SUBAPPLICATION Button_Toggle_RPC_TO_Remote_BG_Option_OPC (* Wie Button_Toggle_RPC_TO_Remote_BG_OPC (IO-Diag-Taster, Loslassen ruft per CLIENT_0 eine RPC-Toggle-Methode auf dem Zielmodul auf, Hintergrundfarbe aus Remote-Subscribe), aber per AOption aktiviert statt QI/INIT. AOption_OUT reicht die Aktivierung nach dem eigenen INIT weiter (Daisy-Chain). *)
  (* Standard: 61499-2; Description: Copyright (c) 2026 Meisterschulen am Ostbahnhof This program and the accompanying materials are made available under the terms of the Eclipse Public License 2.0 which is available at https://www.eclipse.org/legal/epl-2.0/ SPDX-License-Identifier: EPL-2.0 *)
  (* Version 1.1, 2026-10-30, Franz Höpfinger, Meisterschulen am Ostbahnhof, Remote-Clients mit Remote_Init_Retry: Kette (und Option-INIT_CNF) wartet nicht mehr auf die Gegenstation, nach INITO- neuer Versuch nach 2 s (forte #1092, sonst 60 s pro fehlendem Node und danach tot). *)
  (* Version 1.0, 2026-10-17, Franz Höpfinger, Meisterschulen am Ostbahnhof, Kopie von Button_Toggle_RPC_TO_Remote_BG_OPC (Franz: 'kopieren, Variante mit AOption machen') - INIT/INITO/QI/QO ersetzt durch AOption_IN (AOption_X_TO_EVENT) und AOption_OUT (AOption_EVENT_TO_X, Daisy-Chain wie OptionalGroup_001a). AOption_OUT muss weiterverbunden sein (DummyGroup als Kettenende), sonst kommt kein INIT_CNF zurueck. *)
  PACKAGE MyLib::sys;
  IMPORT isobus::UT::Q::const::IDs::ID_NULL;
  IMPORT isobus::UT::io::Button::ButtonActivationCode::BT_RELEASED_UNLATCHED;
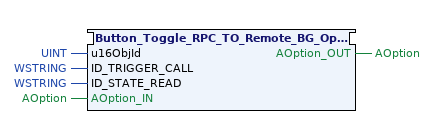
  VAR_INPUT
    u16ObjId : UINT := ID_NULL; (* Object ID Button/Background *)
    ID_TRIGGER_CALL : WSTRING; (* Remote-Methodenadresse (ACTION=CALL_METHOD) fuer den argumentlosen Trigger-Methodenaufruf auf dem Zielmodul *)
    ID_STATE_READ : WSTRING; (* Lokal ueberwachte Adresse (BOOL, ACTION=READ) fuer den Flipflop-Zustand, wird vom Zielmodul remote beschrieben *)
  END_VAR
  SOCKETS
    AOption_IN : Option::AOption; (* Treibt INIT/QI - anschliessen an AOption_AUI_DEMUX_N.OUTx oder AOption_OUT einer vorgeschalteten Instanz *)
  END_SOCKETS
  PLUGS
    AOption_OUT : Option::AOption; (* Reicht die Aktivierung nach dem eigenen INIT an das naechste Glied weiter (Daisy-Chain) - muss verbunden sein, Kettenende z.B. DummyGroup *)
  END_PLUGS
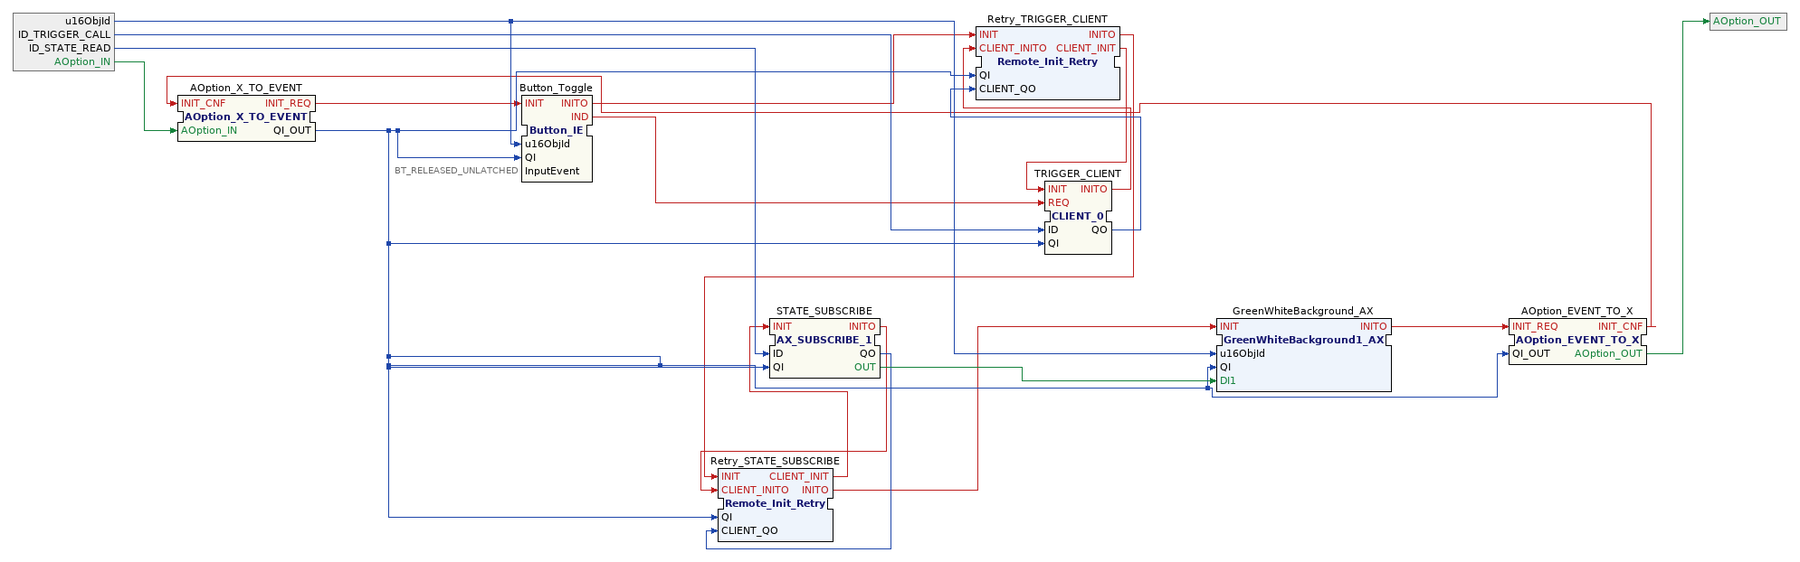
  FBS
    AOption_X_TO_EVENT : Option::conversion::AOption_X_TO_EVENT;
    Button_Toggle : isobus::UT::io::Button::Button_IE(InputEvent := BT_RELEASED_UNLATCHED);
    TRIGGER_CLIENT : iec61499::net::CLIENT_0;
    STATE_SUBSCRIBE : adapter::net::AX_SUBSCRIBE_1;
    AOption_EVENT_TO_X : Option::conversion::AOption_EVENT_TO_X;
  END_FBS
  SUBAPPS
    GreenWhiteBackground_AX : MyLib::sys::GreenWhiteBackground1_AX;
    Retry_TRIGGER_CLIENT : MyLib::sys::Remote_Init_Retry;
    Retry_STATE_SUBSCRIBE : MyLib::sys::Remote_Init_Retry;
  END_SUBAPPS
  EVENT_CONNECTIONS
    Retry_TRIGGER_CLIENT.INITO TO Retry_STATE_SUBSCRIBE.INIT;
    Retry_STATE_SUBSCRIBE.CLIENT_INIT TO STATE_SUBSCRIBE.INIT;
    STATE_SUBSCRIBE.INITO TO Retry_STATE_SUBSCRIBE.CLIENT_INITO;
    Retry_STATE_SUBSCRIBE.INITO TO GreenWhiteBackground_AX.INIT;
    Button_Toggle.INITO TO Retry_TRIGGER_CLIENT.INIT;
    Retry_TRIGGER_CLIENT.CLIENT_INIT TO TRIGGER_CLIENT.INIT;
    TRIGGER_CLIENT.INITO TO Retry_TRIGGER_CLIENT.CLIENT_INITO;
    Button_Toggle.IND TO TRIGGER_CLIENT.REQ;
    AOption_X_TO_EVENT.INIT_REQ TO Button_Toggle.INIT;
    GreenWhiteBackground_AX.INITO TO AOption_EVENT_TO_X.INIT_REQ;
    AOption_EVENT_TO_X.INIT_CNF TO AOption_X_TO_EVENT.INIT_CNF;
  END_CONNECTIONS
  DATA_CONNECTIONS
    AOption_X_TO_EVENT.QI_OUT TO Retry_STATE_SUBSCRIBE.QI;
    STATE_SUBSCRIBE.QO TO Retry_STATE_SUBSCRIBE.CLIENT_QO;
    AOption_X_TO_EVENT.QI_OUT TO Retry_TRIGGER_CLIENT.QI;
    TRIGGER_CLIENT.QO TO Retry_TRIGGER_CLIENT.CLIENT_QO;
    u16ObjId TO Button_Toggle.u16ObjId;
    u16ObjId TO GreenWhiteBackground_AX.u16ObjId;
    ID_TRIGGER_CALL TO TRIGGER_CLIENT.ID;
    ID_STATE_READ TO STATE_SUBSCRIBE.ID;
    AOption_X_TO_EVENT.QI_OUT TO Button_Toggle.QI;
    AOption_X_TO_EVENT.QI_OUT TO TRIGGER_CLIENT.QI;
    AOption_X_TO_EVENT.QI_OUT TO STATE_SUBSCRIBE.QI;
    AOption_X_TO_EVENT.QI_OUT TO GreenWhiteBackground_AX.QI;
    AOption_X_TO_EVENT.QI_OUT TO AOption_EVENT_TO_X.QI_OUT;
  END_CONNECTIONS
  ADAPTER_CONNECTIONS
    AOption_IN TO AOption_X_TO_EVENT.AOption_IN;
    AOption_EVENT_TO_X.AOption_OUT TO AOption_OUT;
    STATE_SUBSCRIBE.OUT TO GreenWhiteBackground_AX.DI1;
  END_CONNECTIONS
END_SUBAPPLICATION
